TYPE ST_EL3356CoeReadData_1 :
STRUCT
	wIdx: WORD;
	bySubIdx: BYTE;
	bReadOK: BOOL;
	dwData: DWORD;
	nSize: UDINT;
END_STRUCT
END_TYPE

(* stored: Version 1.1.0.1, ProductVersion 3.1.4024.15
   DUT ST_EL3356CoeReadData_1: Id {cc215f26-6631-410e-b3f6-146e8e42a296} *)
